% RSLogix 500 project Robot Arm.RSS, saved by version 12.00.00.00 %
PROJECT "SAITO"    % processor: MicroLogix 1400 %

PROGRAM FILES
  LAD 2   38 rungs

DATA FILES
  O0 OUTPUT  7 elements
  I1 INPUT  9 elements
  S2 STATUS  66 elements
  B3 BINARY  16 elements
  T4 TIMER  4 elements
  C5 COUNTER  1 elements
  R6 CONTROL  1 elements
  N7 INTEGER  32 elements
  F8 FLOAT  1 elements
  B13   16 elements
  B14   16 elements

LADDER 2
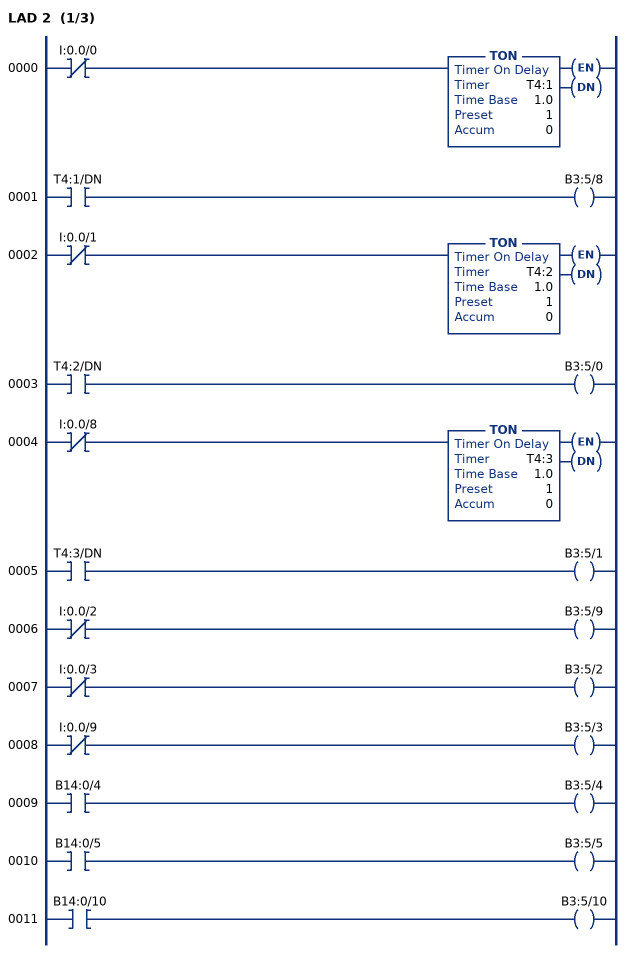
% Rung: 0 %
SOR XIO I:0.0/0 TON T4:1 1.0 1 0 EOR
% Rung: 1 %
SOR XIC T4:1/DN OTE B3:5/8 EOR
% Rung: 2 %
SOR XIO I:0.0/1 TON T4:2 1.0 1 0 EOR
% Rung: 3 %
SOR XIC T4:2/DN OTE B3:5/0 EOR
% Rung: 4 %
SOR XIO I:0.0/8 TON T4:3 1.0 1 0 EOR
% Rung: 5 %
SOR XIC T4:3/DN OTE B3:5/1 EOR
% Rung: 6 %
SOR XIO I:0.0/2 OTE B3:5/9 EOR
% Rung: 7 %
SOR XIO I:0.0/3 OTE B3:5/2 EOR
% Rung: 8 %
SOR XIO I:0.0/9 OTE B3:5/3 EOR
% Rung: 9 %
SOR XIC B14:0/4 OTE B3:5/4 EOR
% Rung: 10 %
SOR XIC B14:0/5 OTE B3:5/5 EOR
% Rung: 11 %
SOR XIC B14:0/10 OTE B3:5/10 EOR

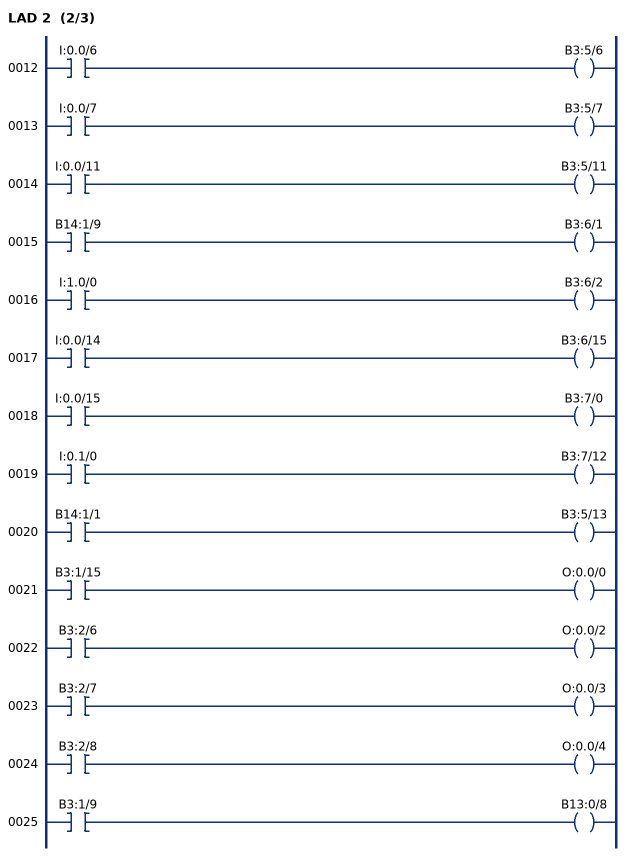
% Rung: 12 %
SOR XIC I:0.0/6 OTE B3:5/6 EOR
% Rung: 13 %
SOR XIC I:0.0/7 OTE B3:5/7 EOR
% Rung: 14 %
SOR XIC I:0.0/11 OTE B3:5/11 EOR
% Rung: 15 %
SOR XIC B14:1/9 OTE B3:6/1 EOR
% Rung: 16 %
SOR XIC I:1.0/0 OTE B3:6/2 EOR
% Rung: 17 %
SOR XIC I:0.0/14 OTE B3:6/15 EOR
% Rung: 18 %
SOR XIC I:0.0/15 OTE B3:7/0 EOR
% Rung: 19 %
SOR XIC I:0.1/0 OTE B3:7/12 EOR
% Rung: 20 %
SOR XIC B14:1/1 OTE B3:5/13 EOR
% Rung: 21 %
SOR XIC B3:1/15 OTE O:0.0/0 EOR
% Rung: 22 %
SOR XIC B3:2/6 OTE O:0.0/2 EOR
% Rung: 23 %
SOR XIC B3:2/7 OTE O:0.0/3 EOR
% Rung: 24 %
SOR XIC B3:2/8 OTE O:0.0/4 EOR
% Rung: 25 %
SOR XIC B3:1/9 OTE B13:0/8 EOR

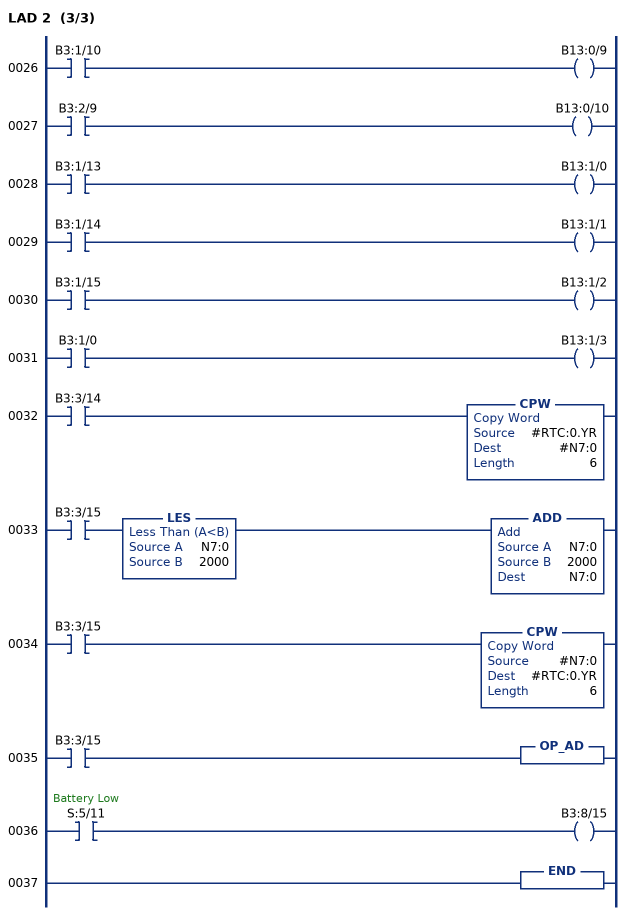
% Rung: 26 %
SOR XIC B3:1/10 OTE B13:0/9 EOR
% Rung: 27 %
SOR XIC B3:2/9 OTE B13:0/10 EOR
% Rung: 28 %
SOR XIC B3:1/13 OTE B13:1/0 EOR
% Rung: 29 %
SOR XIC B3:1/14 OTE B13:1/1 EOR
% Rung: 30 %
SOR XIC B3:1/15 OTE B13:1/2 EOR
% Rung: 31 %
SOR XIC B3:1/0 OTE B13:1/3 EOR
% Rung: 32 %
SOR XIC B3:3/14 CPW #RTC:0.YR #N7:0 6 EOR
% Rung: 33 %
SOR XIC B3:3/15 LES N7:0 2000 ADD N7:0 2000 N7:0 EOR
% Rung: 34 %
SOR XIC B3:3/15 CPW #N7:0 #RTC:0.YR 6 EOR
% Rung: 35 %
SOR XIC B3:3/15 OP_AD EOR
% Rung: 36 %
SOR XIC S:5/11 OTE B3:8/15 EOR
%   S:5/11  "Battery Low" %
% Rung: 37 %
SOR END EOR

DATA TABLE (non-zero values as saved)
DATA B3
% B3:0 % 0X41A7 0X4080 0X0000 0X4000 0X0000 0X220C 0X0000 0X0000 0X0000 0X0000
DATA T4
% .PRE .ACC %
% T4:1 % 1 0
% T4:2 % 1 0
% T4:3 % 1 0
DATA N7
% N7:0 % 2026 10 27 9 1 26 0 0 0 0
DATA B13
% B13:0 % 0X0000 0X0002 0X0000 0X0000 0X0000 0X0000 0X0000 0X0000 0X0000 0X0000
DATA B14
% B14:0 % 0X0000 0X0002 0X0000 0X0000 0X0000 0X0000 0X0000 0X0000 0X0000 0X0000
